// TIA Portal project "MT_SLP333D-IOL_v2" (V18)

(* hardware
DEVICE "S71500/ET200MP station_1"  S7-1500 station
   slot 0: "Rail_0"  Rack  6ES7 590-1***0-0AA0
   slot 1: "PLC_1"  CPU 1516-3 PN/DP  6ES7 516-3AN01-0AB0  V2.8
      slot 3: "CPU display_1"  6ES7591-1BA00-0AA0
      slot 32768: "PROFINET interface_1"  X1
         slot 32769: "Port_1"  X1 P1
         slot 32770: "Port_2"  X1 P2
      slot 33024: "PROFINET interface_2"  X2
         slot 33025: "Port_1"  X2 P1
      slot 33280: "DP interface_1"  X3
      slot 34817: "Virtual CP interface port_1"  Virtual CP interface port  Virtual CP interface port
DEVICE "GSD device_1"  GSD.Device.PN
   slot 0: "Rack"  Rack  V1.0
   slot 0: "bnixg35080b5r067"  BNI XG3-508-0B5-R067  BNI00L3  V1.4.0
      slot 0: "BNI XG3-508-0B5-R067"  BNI XG3-508-0B5-R067
      slot 1: "PN-IO"  PN-IO
         slot 1: "Port XF1"  Port XF1
         slot 2: "Port XF2"  Port XF2
   slot 1: "IO-Link I/O Ports_1"  IO-Link I/O Ports
      slot 0: "BALLUFF 8 Port IO-Link Master"  BALLUFF 8 Port IO-Link Master
   slot 1: "Port deactivated"  Port deactivated
   slot 2: "Port deactivated_1"  Port deactivated
   slot 3: "Port deactivated_2"  Port deactivated
   slot 4: "SLP333D-IOL_Port4I"  IOL_I/O_08/08_Byte + PQI
   slot 5: "Port deactivated_4"  Port deactivated
   slot 6: "Port deactivated_5"  Port deactivated
   slot 7: "Port deactivated_6"  Port deactivated
   slot 8: "Port deactivated_7"  Port deactivated
*)

// ===== PLC "PLC_1"  CPU 1516-3 PN/DP =====

VAR_GLOBAL   // PLC tag table "Default tag table"
   "FirstScan" AT %M1.0 : Bool;
   "SLP/SWP33x_In_Octet0_3" AT %ID1 : DWord;
   "SLP/SWP33x_In_Octet4" AT %IB5 : Byte;
   "SLP/SWP33x_In_Octet5" AT %IB6 : Byte;
   "SLP/SWP33x_In_Octet6" AT %IB7 : Byte;
   "CurrentWeight" AT %MD68 : Real;
   "LowerThreshold" AT %MW72 : UInt;
   "AcyclicCommandIndex" AT %MW74 : UInt;
   "Write_LowerTreshold" AT %M76.0 : Bool;
   "Read_SensorStatus" AT %M76.1 : Bool;
   "Read_AcyclicCommand" AT %M76.2 : Bool;
   "Read_LowerTreshold" AT %M76.3 : Bool;
   "Send_System_Command" AT %M76.4 : Bool;
   "SystemCommand" AT %MW78 : UInt;
   "AcyclicCommandSubindex" AT %MW80 : UInt;
   "AcyclicCommandLength" AT %MW82 : UInt;
   "SensorStatus_SensorNr" AT %MW84 : UInt;
   "Reset_Acyclic_Block" AT %M86.0 : Bool;
   "Smart5Lvl2" AT %M86.1 : Bool;
   "Smart5Lvl3" AT %M86.2 : Bool;
   "Smart5Lvl4" AT %M86.3 : Bool;
   "Smart5Lvl5" AT %M86.4 : Bool;
   "LowerLvlAlarm" AT %M86.5 : Bool;
   "UpperLvlAlarm" AT %M86.6 : Bool;
   "Heartbeat" AT %M86.7 : Bool;
   "CurrentWeightPercent" AT %MD87 : Real;
   "SLP/SWP33x_In_Octet7" AT %IB8 : Byte;
   "SLP/SWP33x_Out_Octet0_3" AT %QD1 : DWord;
   "SLP/SWP33x_Out_Octet6_7" AT %QW7 : Int;
   "ResetCommand" AT %M0.0 : Bool;
   "CommandValue" AT %MD10 : Real;
   "Command" AT %MW15 : Int;
   "WeightMode" AT %MW18 : Int;
   "ProcessType" AT %MW20 : Int;
   "ProcessStatus" AT %MW22 : Int;
   "Write_CommandWithParameter" AT %M76.5 : Bool;
   "ParameterValue" AT %MW91 : UInt;
END_VAR

TYPE "SAI_MB_DeviceStatus"
VERSION : 0.1
   STRUCT
      "Number of Sensors bit 1" : Byte;
      "System Status bit 1" : Bool;
      "System Status bit 2" : Bool;
      "System Status bit 3" : Bool;
      "System Status bit 4" : Bool;
   END_STRUCT;
END_TYPE

TYPE "SAI_SB_3rdStatus"
   STRUCT
      "Measure Unit bit 1" : Bool;
      "Measure Unit bit 2" : Bool;
      "Measure Unit bit 3" : Bool;
      "Measure Unit bit 4" : Bool;
      "Measure Type bit 1" : Bool;
      "Measure Type bit 2" : Bool;
      "Lower Alarm Status" : Bool;
      "Upper Alarm Status" : Bool;
   END_STRUCT;
END_TYPE

TYPE "SAI_SB_2ndStatus"
   STRUCT
      "Smart5 level 5" : Bool;
      "Smart5 level 4" : Bool;
      "Smart5 level 3" : Bool;
      "Smart5 level 2" : Bool;
      Hearbeat : Bool;
   END_STRUCT;
END_TYPE

DATA_BLOCK "SLP/SWP331_IOL_DB"   // DB1
{ S7_Optimized_Access := 'TRUE' }
VERSION : 0.1
// stored: InstanceOfName SLP/SWP331_IOL
"SLP/SWP331_IOL"
BEGIN
END_DATA_BLOCK

DATA_BLOCK "IO_LINK_DEVICE_DB"   // DB2
{ S7_Optimized_Access := 'TRUE' }
AUTHOR : SUP_FA
FAMILY : IO-Link
VERSION : 3.0
// stored: InstanceOfName IO_LINK_DEVICE
"IO_LINK_DEVICE"
BEGIN
END_DATA_BLOCK

DATA_BLOCK "SLP/SWP331_IOL_Acyclic_Commands_DB"   // DB3
{ S7_Optimized_Access := 'TRUE' }
VERSION : 0.1
// stored: InstanceOfName SLP/SWP331_IOL_Acyclic_Commands
"SLP/SWP331_IOL_Acyclic_Commands"
BEGIN
END_DATA_BLOCK

DATA_BLOCK "Data_block_IOL"   // DB14
{ S7_Optimized_Access := 'TRUE' }
VERSION : 0.1
   VAR
      Data : Array[0..231] of Byte;
   END_VAR
BEGIN
END_DATA_BLOCK

FUNCTION_BLOCK "SLP/SWP331_IOL"   // FB1, LAD
{ S7_Optimized_Access := 'TRUE' }
VERSION : 0.1
   VAR_INPUT
      "IO-Link_DevicePort" : Int;
      In_Byte0_3_DWord : DWord;
      In_Byte04 : Byte;
      In_Byte05 : Byte;
      In_Byte06 : Byte;
      In_Byte07 : Byte;
   END_VAR
   VAR_OUTPUT
      CurrentWeight : Real;
      WeightType : String;
      WeightUnit : String;
      Data_OK : Bool;
      Center_Of_Zero : Bool;
      Motion : Bool;
      Net_Mode : Bool;
      Status_Smart5_Lvl_2 : Bool;
      Status_Smart5_Lvl_3 : Bool;
      Status_Smart5_Lvl_4 : Bool;
      Status_Smart5_Lvl_5 : Bool;
      Status_HeartBeat : Bool;
      "Factory adjustment active" : Bool;
      "Last Adjustment Status" : Bool;
      ProcessType : String;
      ProcessType_1 : Int;
      NewWeightUpdate : Bool;
      ProcessStatus : String;
      ProcessStatus_1 : Int;
      Out_Byte0_3_DWord : DWord;
      Out_Byte06_7_Int : Int;
   END_VAR
   VAR_IN_OUT
      "Command Value" : Real;
      Command : Int;
   END_VAR
   VAR
      MeasuredWeightType : Byte;
      MeasuredUnit : Byte;
      ProcessTypeParsen : Byte;
      ProcessStatusParsen : Byte;
      CommandExec : Bool;
   END_VAR
BEGIN

REGION Network 1: Assign IO-Link Device Port Number on the IO-Link Master
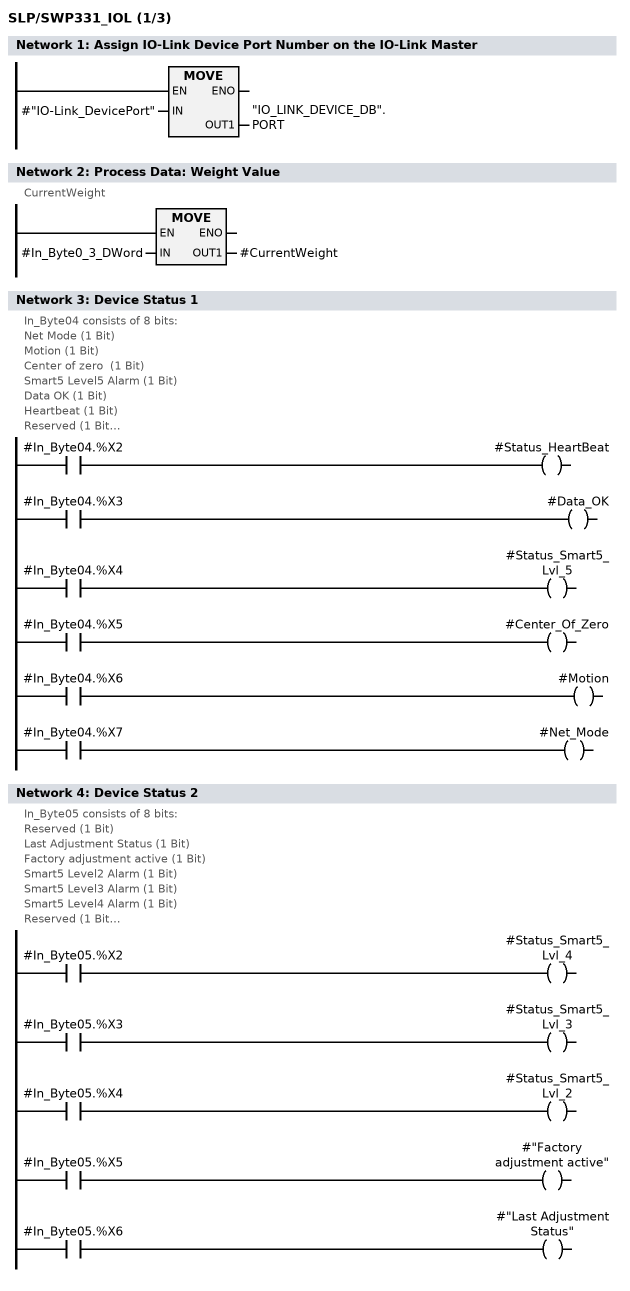
   RUNG wire#powerrail
      Move(in := #"IO-Link_DevicePort", out1 => "IO_LINK_DEVICE_DB".PORT)
   END_RUNG
   // the same network as SCL:
   "IO_LINK_DEVICE_DB".PORT := #"IO-Link_DevicePort";
END_REGION

REGION Network 2: Process Data: Weight Value
   // CurrentWeight
   RUNG wire#powerrail
      Move(in := #In_Byte0_3_DWord, out1 => #CurrentWeight)
   END_RUNG
   // the same network as SCL:
   #CurrentWeight := #In_Byte0_3_DWord;
END_REGION

REGION Network 3: Device Status 1
   // In_Byte04 consists of 8 bits:
   // 
   // Net Mode (1 Bit) 
   // Motion (1 Bit) 
   // Center of zero  (1 Bit) 
   // Smart5 Level5 Alarm (1 Bit) 
   // Data OK (1 Bit) 
   // Heartbeat (1 Bit) 
   // Reserved (1 Bit) 
   // Reserved (1 Bit)
   RUNG wire#powerrail
      Contact( #In_Byte04.%X2 )
      Coil( #Status_HeartBeat )
   END_RUNG
   RUNG wire#powerrail
      Contact( #In_Byte04.%X3 )
      Coil( #Data_OK )
   END_RUNG
   RUNG wire#powerrail
      Contact( #In_Byte04.%X4 )
      Coil( #Status_Smart5_Lvl_5 )
   END_RUNG
   RUNG wire#powerrail
      Contact( #In_Byte04.%X5 )
      Coil( #Center_Of_Zero )
   END_RUNG
   RUNG wire#powerrail
      Contact( #In_Byte04.%X6 )
      Coil( #Motion )
   END_RUNG
   RUNG wire#powerrail
      Contact( #In_Byte04.%X7 )
      Coil( #Net_Mode )
   END_RUNG
   // the same network as SCL:
   #Status_HeartBeat := #In_Byte04.%X2;
   #Data_OK := #In_Byte04.%X3;
   #Status_Smart5_Lvl_5 := #In_Byte04.%X4;
   #Center_Of_Zero := #In_Byte04.%X5;
   #Motion := #In_Byte04.%X6;
   #Net_Mode := #In_Byte04.%X7;
END_REGION

REGION Network 4: Device Status 2
   // In_Byte05 consists of 8 bits:
   // 
   // Reserved (1 Bit) 
   // Last Adjustment Status (1 Bit) 
   // Factory adjustment active (1 Bit) 
   // Smart5 Level2 Alarm (1 Bit)
   // Smart5 Level3 Alarm (1 Bit) 
   // Smart5 Level4 Alarm (1 Bit) 
   // Reserved (1 Bit) 
   // Reserved (1 Bit)
   RUNG wire#powerrail
      Contact( #In_Byte05.%X2 )
      Coil( #Status_Smart5_Lvl_4 )
   END_RUNG
   RUNG wire#powerrail
      Contact( #In_Byte05.%X3 )
      Coil( #Status_Smart5_Lvl_3 )
   END_RUNG
   RUNG wire#powerrail
      Contact( #In_Byte05.%X4 )
      Coil( #Status_Smart5_Lvl_2 )
   END_RUNG
   RUNG wire#powerrail
      Contact( #In_Byte05.%X5 )
      Coil( #"Factory adjustment active" )
   END_RUNG
   RUNG wire#powerrail
      Contact( #In_Byte05.%X6 )
      Coil( #"Last Adjustment Status" )
   END_RUNG
   // the same network as SCL:
   #Status_Smart5_Lvl_4 := #In_Byte05.%X2;
   #Status_Smart5_Lvl_3 := #In_Byte05.%X3;
   #Status_Smart5_Lvl_2 := #In_Byte05.%X4;
   #"Factory adjustment active" := #In_Byte05.%X5;
   #"Last Adjustment Status" := #In_Byte05.%X6;
END_REGION

REGION Network 5: Device Status 3
   // In_Byte06 consists of 8 bits:
   // 
   // Process Type (3 Bit) 
   // New weight update (1 Bit) 
   // Process Status (4 Bit)
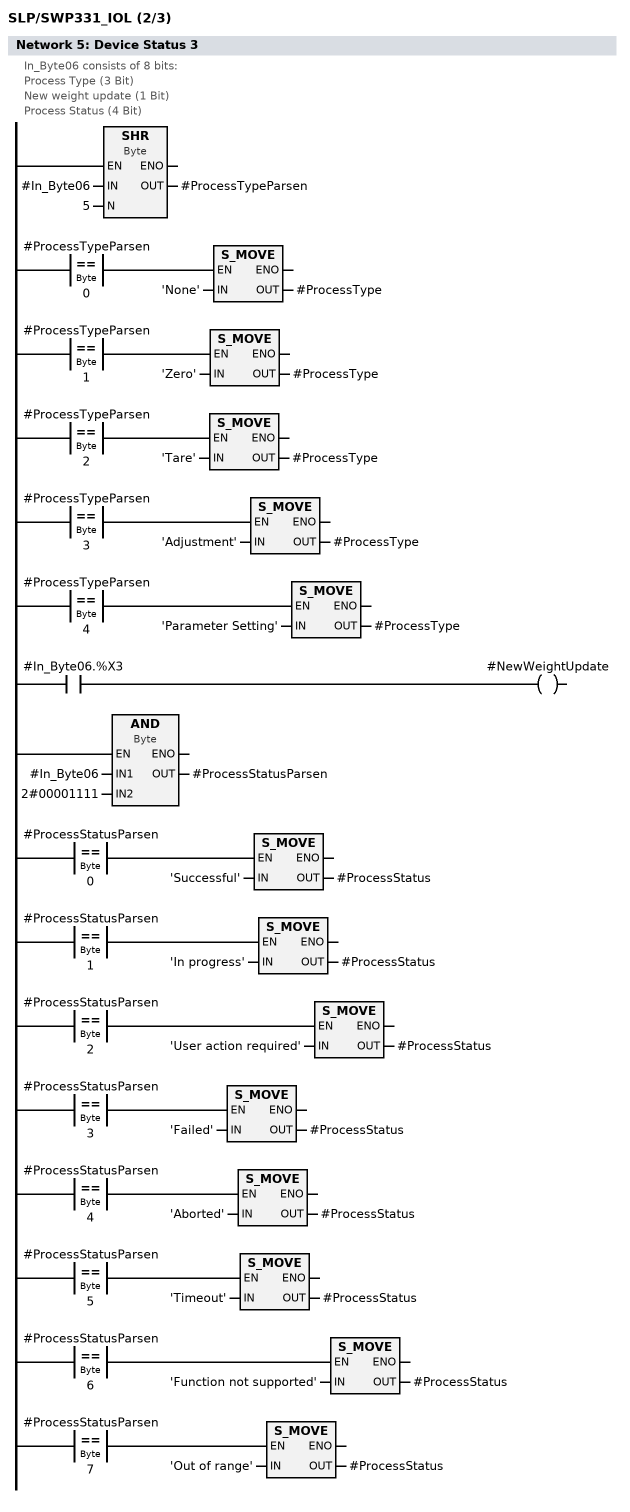
   RUNG wire#powerrail
      { S7_Templates := "SrcType := Byte" } Shr(in := #In_Byte06, n := 5, out => #ProcessTypeParsen)
   END_RUNG
   RUNG wire#powerrail
      { S7_Templates := "SrcType := Byte" } EQ_Contact(in1 := #ProcessTypeParsen, in2 := 0)
      S_Move(in := 'None', out => #ProcessType)
   END_RUNG
   RUNG wire#powerrail
      { S7_Templates := "SrcType := Byte" } EQ_Contact(in1 := #ProcessTypeParsen, in2 := 1)
      S_Move(in := 'Zero', out => #ProcessType)
   END_RUNG
   RUNG wire#powerrail
      { S7_Templates := "SrcType := Byte" } EQ_Contact(in1 := #ProcessTypeParsen, in2 := 2)
      S_Move(in := 'Tare', out => #ProcessType)
   END_RUNG
   RUNG wire#powerrail
      { S7_Templates := "SrcType := Byte" } EQ_Contact(in1 := #ProcessTypeParsen, in2 := 3)
      S_Move(in := 'Adjustment', out => #ProcessType)
   END_RUNG
   RUNG wire#powerrail
      { S7_Templates := "SrcType := Byte" } EQ_Contact(in1 := #ProcessTypeParsen, in2 := 4)
      S_Move(in := 'Parameter Setting', out => #ProcessType)
   END_RUNG
   RUNG wire#powerrail
      Contact( #In_Byte06.%X3 )
      Coil( #NewWeightUpdate )
   END_RUNG
   RUNG wire#powerrail
      { S7_Templates := "SrcType := Byte" } And(in1 := #In_Byte06, in2 := 2#00001111, out => #ProcessStatusParsen)
   END_RUNG
   RUNG wire#powerrail
      { S7_Templates := "SrcType := Byte" } EQ_Contact(in1 := #ProcessStatusParsen, in2 := 0)
      S_Move(in := 'Successful', out => #ProcessStatus)
   END_RUNG
   RUNG wire#powerrail
      { S7_Templates := "SrcType := Byte" } EQ_Contact(in1 := #ProcessStatusParsen, in2 := 1)
      S_Move(in := 'In progress', out => #ProcessStatus)
   END_RUNG
   RUNG wire#powerrail
      { S7_Templates := "SrcType := Byte" } EQ_Contact(in1 := #ProcessStatusParsen, in2 := 2)
      S_Move(in := 'User action required', out => #ProcessStatus)
   END_RUNG
   RUNG wire#powerrail
      { S7_Templates := "SrcType := Byte" } EQ_Contact(in1 := #ProcessStatusParsen, in2 := 3)
      S_Move(in := 'Failed', out => #ProcessStatus)
   END_RUNG
   RUNG wire#powerrail
      { S7_Templates := "SrcType := Byte" } EQ_Contact(in1 := #ProcessStatusParsen, in2 := 4)
      S_Move(in := 'Aborted', out => #ProcessStatus)
   END_RUNG
   RUNG wire#powerrail
      { S7_Templates := "SrcType := Byte" } EQ_Contact(in1 := #ProcessStatusParsen, in2 := 5)
      S_Move(in := 'Timeout', out => #ProcessStatus)
   END_RUNG
   RUNG wire#powerrail
      { S7_Templates := "SrcType := Byte" } EQ_Contact(in1 := #ProcessStatusParsen, in2 := 6)
      S_Move(in := 'Function not supported', out => #ProcessStatus)
   END_RUNG
   RUNG wire#powerrail
      { S7_Templates := "SrcType := Byte" } EQ_Contact(in1 := #ProcessStatusParsen, in2 := 7)
      S_Move(in := 'Out of range', out => #ProcessStatus)
   END_RUNG
   // the same network as SCL:
   #ProcessTypeParsen := SHR(IN := #In_Byte06, N := 5);
   IF #ProcessTypeParsen = 0 THEN #ProcessType := 'None'; END_IF;
   IF #ProcessTypeParsen = 1 THEN #ProcessType := 'Zero'; END_IF;
   IF #ProcessTypeParsen = 2 THEN #ProcessType := 'Tare'; END_IF;
   IF #ProcessTypeParsen = 3 THEN #ProcessType := 'Adjustment'; END_IF;
   IF #ProcessTypeParsen = 4 THEN #ProcessType := 'Parameter Setting'; END_IF;
   #NewWeightUpdate := #In_Byte06.%X3;
   #ProcessStatusParsen := #In_Byte06 AND 2#00001111;
   IF #ProcessStatusParsen = 0 THEN #ProcessStatus := 'Successful'; END_IF;
   IF #ProcessStatusParsen = 1 THEN #ProcessStatus := 'In progress'; END_IF;
   IF #ProcessStatusParsen = 2 THEN #ProcessStatus := 'User action required'; END_IF;
   IF #ProcessStatusParsen = 3 THEN #ProcessStatus := 'Failed'; END_IF;
   IF #ProcessStatusParsen = 4 THEN #ProcessStatus := 'Aborted'; END_IF;
   IF #ProcessStatusParsen = 5 THEN #ProcessStatus := 'Timeout'; END_IF;
   IF #ProcessStatusParsen = 6 THEN #ProcessStatus := 'Function not supported'; END_IF;
   IF #ProcessStatusParsen = 7 THEN #ProcessStatus := 'Out of range'; END_IF;
END_REGION

REGION Network 6: Weight Information
   // In_Byte07 consists of 8 bits:
   // Weight Type (4 Bits)
   // Weight Unit (4 Bits)
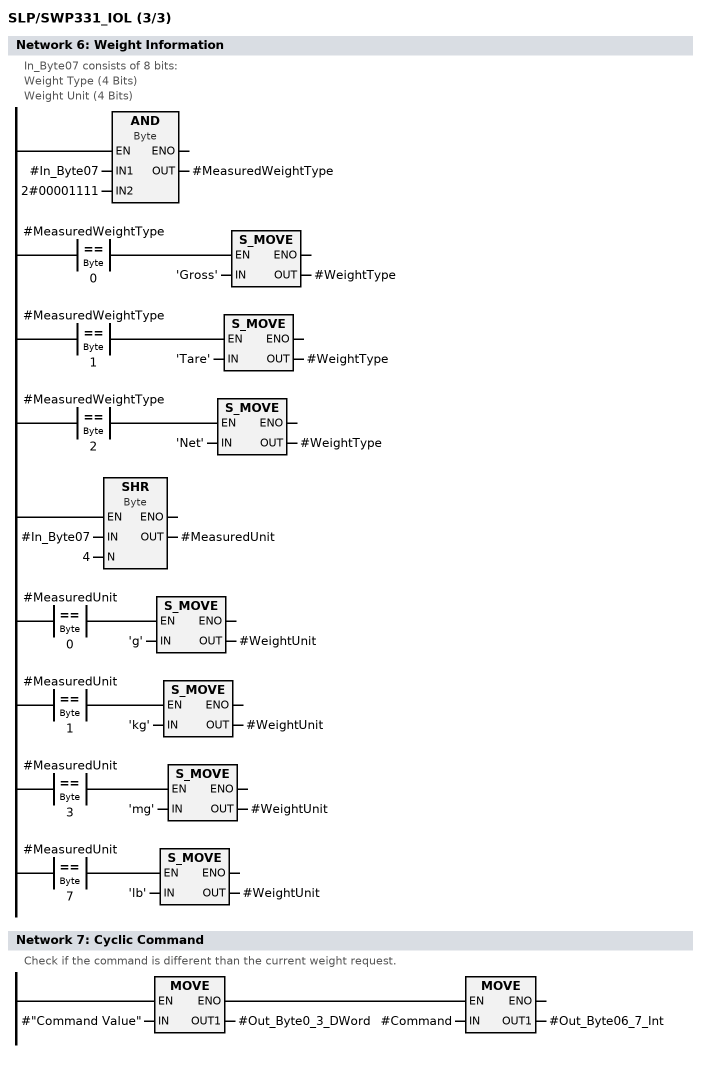
   RUNG wire#powerrail
      { S7_Templates := "SrcType := Byte" } And(in1 := #In_Byte07, in2 := 2#00001111, out => #MeasuredWeightType)
   END_RUNG
   RUNG wire#powerrail
      { S7_Templates := "SrcType := Byte" } EQ_Contact(in1 := #MeasuredWeightType, in2 := 0)
      S_Move(in := 'Gross', out => #WeightType)
   END_RUNG
   RUNG wire#powerrail
      { S7_Templates := "SrcType := Byte" } EQ_Contact(in1 := #MeasuredWeightType, in2 := 1)
      S_Move(in := 'Tare', out => #WeightType)
   END_RUNG
   RUNG wire#powerrail
      { S7_Templates := "SrcType := Byte" } EQ_Contact(in1 := #MeasuredWeightType, in2 := 2)
      S_Move(in := 'Net', out => #WeightType)
   END_RUNG
   RUNG wire#powerrail
      { S7_Templates := "SrcType := Byte" } Shr(in := #In_Byte07, n := 4, out => #MeasuredUnit)
   END_RUNG
   RUNG wire#powerrail
      { S7_Templates := "SrcType := Byte" } EQ_Contact(in1 := #MeasuredUnit, in2 := 0)
      S_Move(in := 'g', out => #WeightUnit)
   END_RUNG
   RUNG wire#powerrail
      { S7_Templates := "SrcType := Byte" } EQ_Contact(in1 := #MeasuredUnit, in2 := 1)
      S_Move(in := 'kg', out => #WeightUnit)
   END_RUNG
   RUNG wire#powerrail
      { S7_Templates := "SrcType := Byte" } EQ_Contact(in1 := #MeasuredUnit, in2 := 3)
      S_Move(in := 'mg', out => #WeightUnit)
   END_RUNG
   RUNG wire#powerrail
      { S7_Templates := "SrcType := Byte" } EQ_Contact(in1 := #MeasuredUnit, in2 := 7)
      S_Move(in := 'lb', out => #WeightUnit)
   END_RUNG
   // the same network as SCL:
   #MeasuredWeightType := #In_Byte07 AND 2#00001111;
   IF #MeasuredWeightType = 0 THEN #WeightType := 'Gross'; END_IF;
   IF #MeasuredWeightType = 1 THEN #WeightType := 'Tare'; END_IF;
   IF #MeasuredWeightType = 2 THEN #WeightType := 'Net'; END_IF;
   #MeasuredUnit := SHR(IN := #In_Byte07, N := 4);
   IF #MeasuredUnit = 0 THEN #WeightUnit := 'g'; END_IF;
   IF #MeasuredUnit = 1 THEN #WeightUnit := 'kg'; END_IF;
   IF #MeasuredUnit = 3 THEN #WeightUnit := 'mg'; END_IF;
   IF #MeasuredUnit = 7 THEN #WeightUnit := 'lb'; END_IF;
END_REGION

REGION Network 7: Cyclic Command
   // Check if the command is different than the current weight request.
   RUNG wire#powerrail
      Move(in := #"Command Value", out1 => #Out_Byte0_3_DWord)
      Move(in := #Command, out1 => #Out_Byte06_7_Int)
   END_RUNG
   // the same network as SCL:
   #Out_Byte0_3_DWord := #"Command Value";
   #Out_Byte06_7_Int := #Command;
END_REGION
END_FUNCTION_BLOCK

FUNCTION_BLOCK "SLP/SWP331_IOL_Acyclic_Commands"   // FB2, LAD
{ S7_Optimized_Access := 'TRUE' }
VERSION : 0.1
   VAR_INPUT
      SystemCommand : UInt;
      AcyclicCommandIndex : UInt;
      AcyclicCommandSubindex : UInt;
      AcyclicCommandLength : UInt;
      ParameterValue : UInt;
   END_VAR
   VAR_OUTPUT
      SensorStatus : Byte;
      ErrorCode : DWord;
      Done : Bool;
   END_VAR
   VAR_IN_OUT
      Send_SystemCmd : Bool;
      Write_AcyclicCommandWithParameter : Bool;
      Read_AcyclicCommand : Bool;
      ResetAcyclicBlock : Bool;
   END_VAR
   VAR
      WriteStep : SInt;
      ReadStep : SInt;
      Cmd_RWTrigger : Bool;
   END_VAR
   VAR_TEMP   // added for the SCL form of the ladder/FBD networks
      _w1 : Bool;
      _w2 : Bool;
      _w3 : Bool;
      _w4 : Bool;
      _w5 : Bool;
      _w6 : Bool;
   END_VAR
BEGIN

REGION Network 1: Send Acyclic Command
   // Change the variable #SystemCommand in the Application Block and trigger the #Send_SystemCmd to send a system command to the device.
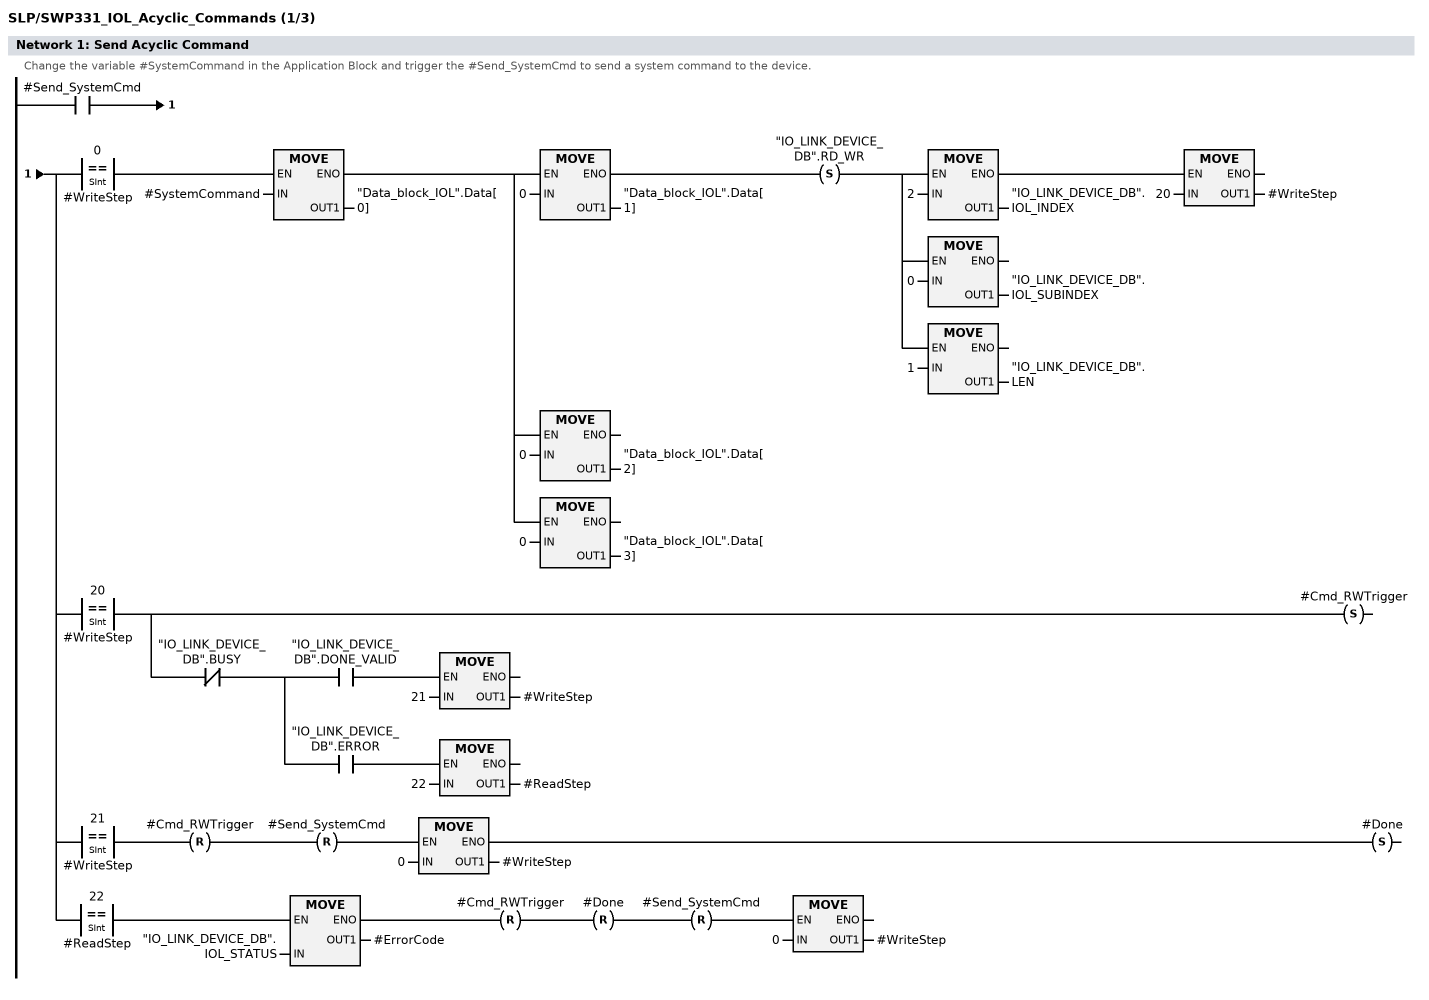
   RUNG wire#powerrail
      Contact( #Send_SystemCmd )
      wire#w1
      { S7_Templates := "SrcType := SInt" } EQ_Contact(in1 := 0, in2 := #WriteStep)
      Move(in := #SystemCommand, out1 => "Data_block_IOL".Data[0])
      wire#w2
      Move(in := 0, out1 => "Data_block_IOL".Data[1])
      S_Coil( "IO_LINK_DEVICE_DB".RD_WR )
      wire#w3
      Move(in := 2, out1 => "IO_LINK_DEVICE_DB".IOL_INDEX)
      Move(in := 20, out1 => #WriteStep)
   END_RUNG
   RUNG wire#w3
      Move(in := 0, out1 => "IO_LINK_DEVICE_DB".IOL_SUBINDEX)
   END_RUNG
   RUNG wire#w3
      Move(in := 1, out1 => "IO_LINK_DEVICE_DB".LEN)
   END_RUNG
   RUNG wire#w2
      Move(in := 0, out1 => "Data_block_IOL".Data[2])
   END_RUNG
   RUNG wire#w2
      Move(in := 0, out1 => "Data_block_IOL".Data[3])
   END_RUNG
   RUNG wire#w1
      { S7_Templates := "SrcType := SInt" } EQ_Contact(in1 := 20, in2 := #WriteStep)
      wire#w4
      S_Coil( #Cmd_RWTrigger )
   END_RUNG
   RUNG wire#w4
      I_Contact( "IO_LINK_DEVICE_DB".BUSY )
      wire#w5
      Contact( "IO_LINK_DEVICE_DB".DONE_VALID )
      Move(in := 21, out1 => #WriteStep)
   END_RUNG
   RUNG wire#w5
      Contact( "IO_LINK_DEVICE_DB".ERROR )
      Move(in := 22, out1 => #ReadStep)
   END_RUNG
   RUNG wire#w1
      { S7_Templates := "SrcType := SInt" } EQ_Contact(in1 := 21, in2 := #WriteStep)
      R_Coil( #Cmd_RWTrigger )
      R_Coil( #Send_SystemCmd )
      Move(in := 0, out1 => #WriteStep)
      S_Coil( #Done )
   END_RUNG
   RUNG wire#w1
      { S7_Templates := "SrcType := SInt" } EQ_Contact(in1 := 22, in2 := #ReadStep)
      Move(in := "IO_LINK_DEVICE_DB".IOL_STATUS, out1 => #ErrorCode)
      R_Coil( #Cmd_RWTrigger )
      R_Coil( #Done )
      R_Coil( #Send_SystemCmd )
      Move(in := 0, out1 => #WriteStep)
   END_RUNG
   // the same network as SCL:
   IF #Send_SystemCmd AND (0 = #WriteStep) THEN
       "Data_block_IOL".Data[0] := #SystemCommand;
       "Data_block_IOL".Data[1] := 0;
       "IO_LINK_DEVICE_DB".RD_WR := TRUE;
       "IO_LINK_DEVICE_DB".IOL_INDEX := 2;
   END_IF;
   #_w1 := #Send_SystemCmd AND (0 = #WriteStep);
   #_w2 := #Send_SystemCmd AND (0 = #WriteStep);
   IF #_w2 THEN
       #WriteStep := 20;
       "IO_LINK_DEVICE_DB".IOL_SUBINDEX := 0;
       "IO_LINK_DEVICE_DB".LEN := 1;
   END_IF;
   IF #_w1 THEN
       "Data_block_IOL".Data[2] := 0;
       "Data_block_IOL".Data[3] := 0;
   END_IF;
   #_w3 := #Send_SystemCmd AND (20 = #WriteStep);
   IF #_w3 THEN #Cmd_RWTrigger := TRUE; END_IF;
   #_w4 := #_w3 AND NOT "IO_LINK_DEVICE_DB".BUSY;
   IF #_w4 AND "IO_LINK_DEVICE_DB".DONE_VALID THEN #WriteStep := 21; END_IF;
   IF #_w4 AND "IO_LINK_DEVICE_DB".ERROR THEN #ReadStep := 22; END_IF;
   IF #Send_SystemCmd AND (21 = #WriteStep) THEN #Cmd_RWTrigger := FALSE; END_IF;
   #_w5 := #Send_SystemCmd AND (21 = #WriteStep);
   #_w6 := #Send_SystemCmd;
   IF #_w5 THEN
       #Send_SystemCmd := FALSE;
       #WriteStep := 0;
       #Done := TRUE;
   END_IF;
   IF #_w6 AND (22 = #ReadStep) THEN
       #ErrorCode := "IO_LINK_DEVICE_DB".IOL_STATUS;
       #Cmd_RWTrigger := FALSE;
       #Done := FALSE;
       #Send_SystemCmd := FALSE;
       #WriteStep := 0;
   END_IF;
END_REGION

REGION Network 2: Read Acyclic Command
   // Change the variables value #AcyclicCommandIndex, #AcyclicCommandSubindex and #AcyclicCommandLength in the Application Block and trigger the #Read_AcyclicCommand to send an acyclic command to the device.
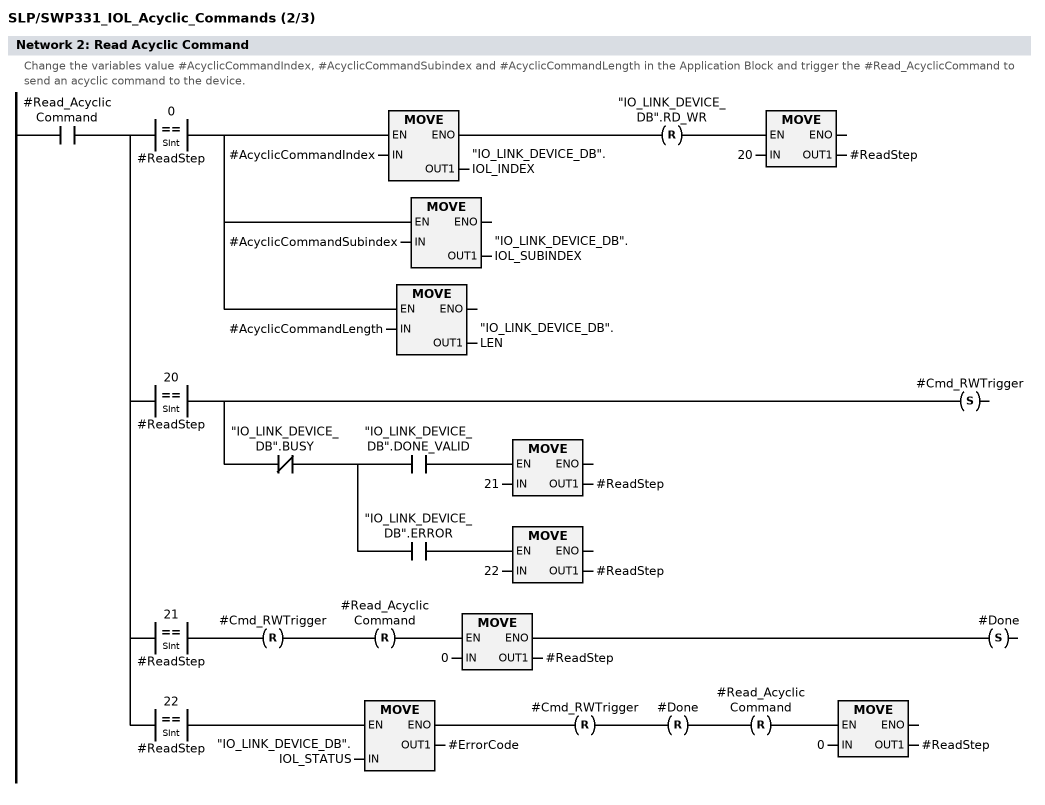
   RUNG wire#powerrail
      Contact( #Read_AcyclicCommand )
      wire#w1
      { S7_Templates := "SrcType := SInt" } EQ_Contact(in1 := 0, in2 := #ReadStep)
      wire#w2
      Move(in := #AcyclicCommandIndex, out1 => "IO_LINK_DEVICE_DB".IOL_INDEX)
      R_Coil( "IO_LINK_DEVICE_DB".RD_WR )
      Move(in := 20, out1 => #ReadStep)
   END_RUNG
   RUNG wire#w2
      Move(in := #AcyclicCommandSubindex, out1 => "IO_LINK_DEVICE_DB".IOL_SUBINDEX)
   END_RUNG
   RUNG wire#w2
      Move(in := #AcyclicCommandLength, out1 => "IO_LINK_DEVICE_DB".LEN)
   END_RUNG
   RUNG wire#w1
      { S7_Templates := "SrcType := SInt" } EQ_Contact(in1 := 20, in2 := #ReadStep)
      wire#w3
      S_Coil( #Cmd_RWTrigger )
   END_RUNG
   RUNG wire#w3
      I_Contact( "IO_LINK_DEVICE_DB".BUSY )
      wire#w4
      Contact( "IO_LINK_DEVICE_DB".DONE_VALID )
      Move(in := 21, out1 => #ReadStep)
   END_RUNG
   RUNG wire#w4
      Contact( "IO_LINK_DEVICE_DB".ERROR )
      Move(in := 22, out1 => #ReadStep)
   END_RUNG
   RUNG wire#w1
      { S7_Templates := "SrcType := SInt" } EQ_Contact(in1 := 21, in2 := #ReadStep)
      R_Coil( #Cmd_RWTrigger )
      R_Coil( #Read_AcyclicCommand )
      Move(in := 0, out1 => #ReadStep)
      S_Coil( #Done )
   END_RUNG
   RUNG wire#w1
      { S7_Templates := "SrcType := SInt" } EQ_Contact(in1 := 22, in2 := #ReadStep)
      Move(in := "IO_LINK_DEVICE_DB".IOL_STATUS, out1 => #ErrorCode)
      R_Coil( #Cmd_RWTrigger )
      R_Coil( #Done )
      R_Coil( #Read_AcyclicCommand )
      Move(in := 0, out1 => #ReadStep)
   END_RUNG
   // the same network as SCL:
   IF #Read_AcyclicCommand AND (0 = #ReadStep) THEN
       "IO_LINK_DEVICE_DB".IOL_INDEX := #AcyclicCommandIndex;
       "IO_LINK_DEVICE_DB".RD_WR := FALSE;
   END_IF;
   #_w1 := #Read_AcyclicCommand AND (0 = #ReadStep);
   IF #_w1 THEN
       #ReadStep := 20;
       "IO_LINK_DEVICE_DB".IOL_SUBINDEX := #AcyclicCommandSubindex;
       "IO_LINK_DEVICE_DB".LEN := #AcyclicCommandLength;
   END_IF;
   #_w2 := #Read_AcyclicCommand AND (20 = #ReadStep);
   IF #_w2 THEN #Cmd_RWTrigger := TRUE; END_IF;
   #_w3 := #_w2 AND NOT "IO_LINK_DEVICE_DB".BUSY;
   IF #_w3 AND "IO_LINK_DEVICE_DB".DONE_VALID THEN #ReadStep := 21; END_IF;
   IF #_w3 AND "IO_LINK_DEVICE_DB".ERROR THEN #ReadStep := 22; END_IF;
   IF #Read_AcyclicCommand AND (21 = #ReadStep) THEN #Cmd_RWTrigger := FALSE; END_IF;
   #_w4 := #Read_AcyclicCommand AND (21 = #ReadStep);
   #_w5 := #Read_AcyclicCommand;
   IF #_w4 THEN
       #Read_AcyclicCommand := FALSE;
       #ReadStep := 0;
       #Done := TRUE;
   END_IF;
   IF #_w5 AND (22 = #ReadStep) THEN
       #ErrorCode := "IO_LINK_DEVICE_DB".IOL_STATUS;
       #Cmd_RWTrigger := FALSE;
       #Done := FALSE;
       #Read_AcyclicCommand := FALSE;
       #ReadStep := 0;
   END_IF;
END_REGION

REGION Network 3: Write Acyclic Command
   // Change the variables value #AcyclicCommandIndex, #AcyclicCommandSubindex #ParameterValue and #AcyclicCommandLength in the Application Block and trigger the #Write_AcyclicCommand to send an acyclic command to the device.
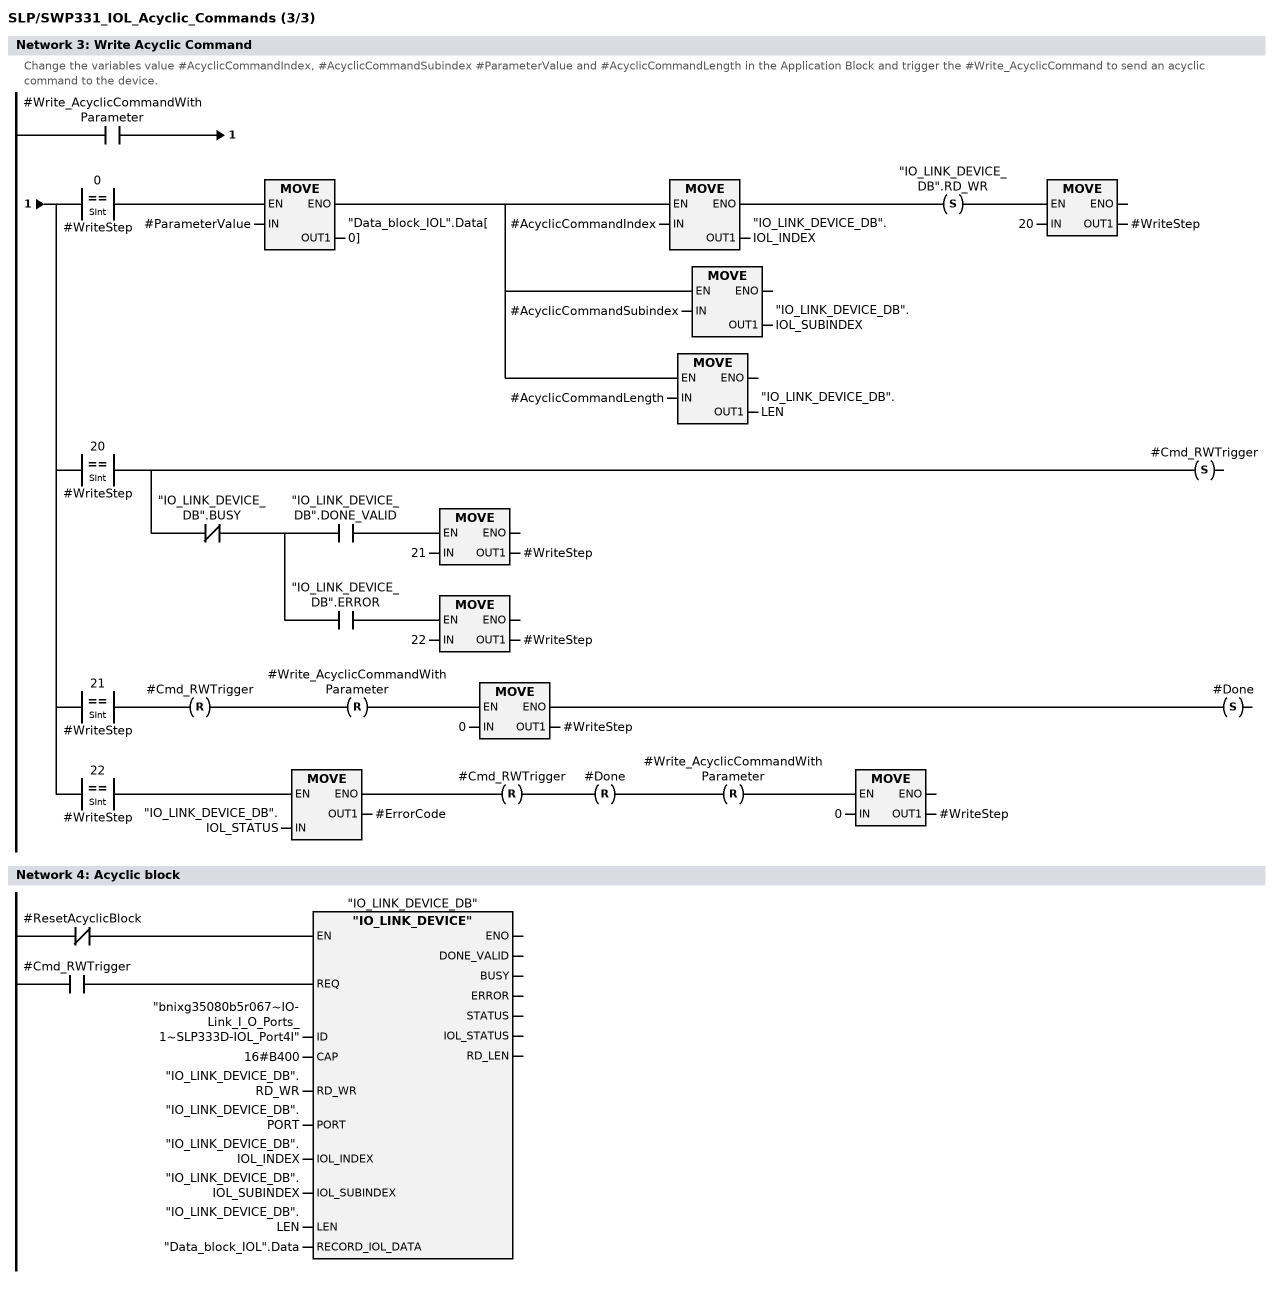
   RUNG wire#powerrail
      Contact( #Write_AcyclicCommandWithParameter )
      wire#w1
      { S7_Templates := "SrcType := SInt" } EQ_Contact(in1 := 0, in2 := #WriteStep)
      Move(in := #ParameterValue, out1 => "Data_block_IOL".Data[0])
      wire#w2
      Move(in := #AcyclicCommandIndex, out1 => "IO_LINK_DEVICE_DB".IOL_INDEX)
      S_Coil( "IO_LINK_DEVICE_DB".RD_WR )
      Move(in := 20, out1 => #WriteStep)
   END_RUNG
   RUNG wire#w2
      Move(in := #AcyclicCommandSubindex, out1 => "IO_LINK_DEVICE_DB".IOL_SUBINDEX)
   END_RUNG
   RUNG wire#w2
      Move(in := #AcyclicCommandLength, out1 => "IO_LINK_DEVICE_DB".LEN)
   END_RUNG
   RUNG wire#w1
      { S7_Templates := "SrcType := SInt" } EQ_Contact(in1 := 20, in2 := #WriteStep)
      wire#w3
      S_Coil( #Cmd_RWTrigger )
   END_RUNG
   RUNG wire#w3
      I_Contact( "IO_LINK_DEVICE_DB".BUSY )
      wire#w4
      Contact( "IO_LINK_DEVICE_DB".DONE_VALID )
      Move(in := 21, out1 => #WriteStep)
   END_RUNG
   RUNG wire#w4
      Contact( "IO_LINK_DEVICE_DB".ERROR )
      Move(in := 22, out1 => #WriteStep)
   END_RUNG
   RUNG wire#w1
      { S7_Templates := "SrcType := SInt" } EQ_Contact(in1 := 21, in2 := #WriteStep)
      R_Coil( #Cmd_RWTrigger )
      R_Coil( #Write_AcyclicCommandWithParameter )
      Move(in := 0, out1 => #WriteStep)
      S_Coil( #Done )
   END_RUNG
   RUNG wire#w1
      { S7_Templates := "SrcType := SInt" } EQ_Contact(in1 := 22, in2 := #WriteStep)
      Move(in := "IO_LINK_DEVICE_DB".IOL_STATUS, out1 => #ErrorCode)
      R_Coil( #Cmd_RWTrigger )
      R_Coil( #Done )
      R_Coil( #Write_AcyclicCommandWithParameter )
      Move(in := 0, out1 => #WriteStep)
   END_RUNG
   // the same network as SCL:
   IF #Write_AcyclicCommandWithParameter AND (0 = #WriteStep) THEN
       "Data_block_IOL".Data[0] := #ParameterValue;
       "IO_LINK_DEVICE_DB".IOL_INDEX := #AcyclicCommandIndex;
       "IO_LINK_DEVICE_DB".RD_WR := TRUE;
   END_IF;
   #_w1 := #Write_AcyclicCommandWithParameter AND (0 = #WriteStep);
   IF #_w1 THEN
       #WriteStep := 20;
       "IO_LINK_DEVICE_DB".IOL_SUBINDEX := #AcyclicCommandSubindex;
       "IO_LINK_DEVICE_DB".LEN := #AcyclicCommandLength;
   END_IF;
   #_w2 := #Write_AcyclicCommandWithParameter AND (20 = #WriteStep);
   IF #_w2 THEN #Cmd_RWTrigger := TRUE; END_IF;
   #_w3 := #_w2 AND NOT "IO_LINK_DEVICE_DB".BUSY;
   IF #_w3 AND "IO_LINK_DEVICE_DB".DONE_VALID THEN #WriteStep := 21; END_IF;
   IF #_w3 AND "IO_LINK_DEVICE_DB".ERROR THEN #WriteStep := 22; END_IF;
   IF #Write_AcyclicCommandWithParameter AND (21 = #WriteStep) THEN #Cmd_RWTrigger := FALSE; END_IF;
   #_w4 := #Write_AcyclicCommandWithParameter AND (21 = #WriteStep);
   #_w5 := #Write_AcyclicCommandWithParameter;
   IF #_w4 THEN
       #Write_AcyclicCommandWithParameter := FALSE;
       #WriteStep := 0;
       #Done := TRUE;
   END_IF;
   IF #_w5 AND (22 = #WriteStep) THEN
       #ErrorCode := "IO_LINK_DEVICE_DB".IOL_STATUS;
       #Cmd_RWTrigger := FALSE;
       #Done := FALSE;
       #Write_AcyclicCommandWithParameter := FALSE;
       #WriteStep := 0;
   END_IF;
END_REGION

REGION Network 4: Acyclic block
   RUNG wire#powerrail
      I_Contact( #ResetAcyclicBlock )
      "IO_LINK_DEVICE_DB"(REQ := wire#w1, ID := "bnixg35080b5r067~IO-Link_I_O_Ports_1~SLP333D-IOL_Port4I", CAP := 16#B400, RD_WR := "IO_LINK_DEVICE_DB".RD_WR, PORT := "IO_LINK_DEVICE_DB".PORT, IOL_INDEX := "IO_LINK_DEVICE_DB".IOL_INDEX, IOL_SUBINDEX := "IO_LINK_DEVICE_DB".IOL_SUBINDEX, LEN := "IO_LINK_DEVICE_DB".LEN, RECORD_IOL_DATA := "Data_block_IOL".Data, DONE_VALID =>, BUSY =>, ERROR =>, STATUS =>, IOL_STATUS =>, RD_LEN =>)
   END_RUNG
   RUNG wire#powerrail
      Contact( #Cmd_RWTrigger )
   END_RUNG wire#w1
   // the same network as SCL:
   IF NOT #ResetAcyclicBlock THEN
       "IO_LINK_DEVICE_DB"(REQ := #Cmd_RWTrigger,   // "IO_LINK_DEVICE"
                           ID := "bnixg35080b5r067~IO-Link_I_O_Ports_1~SLP333D-IOL_Port4I",
                           CAP := 16#B400,
                           RD_WR := "IO_LINK_DEVICE_DB".RD_WR,
                           PORT := "IO_LINK_DEVICE_DB".PORT,
                           IOL_INDEX := "IO_LINK_DEVICE_DB".IOL_INDEX,
                           IOL_SUBINDEX := "IO_LINK_DEVICE_DB".IOL_SUBINDEX,
                           LEN := "IO_LINK_DEVICE_DB".LEN,
                           RECORD_IOL_DATA := "Data_block_IOL".Data);
   END_IF;
END_REGION
END_FUNCTION_BLOCK

FUNCTION "MT_IND_Application" : Void   // FC1, LAD
{ S7_Optimized_Access := 'TRUE' }
VERSION : 0.1
BEGIN

REGION Network 1: Cyclic Data
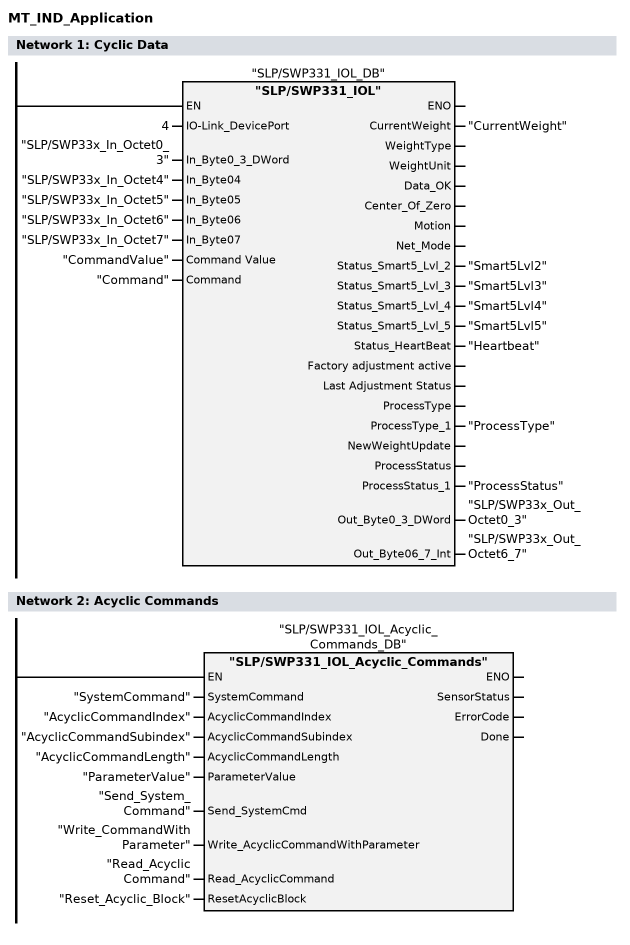
   RUNG wire#powerrail
      "SLP/SWP331_IOL_DB"("IO-Link_DevicePort" := 4, In_Byte0_3_DWord := "SLP/SWP33x_In_Octet0_3", In_Byte04 := "SLP/SWP33x_In_Octet4", In_Byte05 := "SLP/SWP33x_In_Octet5", In_Byte06 := "SLP/SWP33x_In_Octet6", In_Byte07 := "SLP/SWP33x_In_Octet7", "Command Value" := "CommandValue", Command := "Command", CurrentWeight => "CurrentWeight", WeightType =>, WeightUnit =>, Data_OK =>, Center_Of_Zero =>, Motion =>, Net_Mode =>, Status_Smart5_Lvl_2 => "Smart5Lvl2", Status_Smart5_Lvl_3 => "Smart5Lvl3", Status_Smart5_Lvl_4 => "Smart5Lvl4", Status_Smart5_Lvl_5 => "Smart5Lvl5", Status_HeartBeat => "Heartbeat", "Factory adjustment active" =>, "Last Adjustment Status" =>, ProcessType =>, ProcessType_1 => "ProcessType", NewWeightUpdate =>, ProcessStatus =>, ProcessStatus_1 => "ProcessStatus", Out_Byte0_3_DWord => "SLP/SWP33x_Out_Octet0_3", Out_Byte06_7_Int => "SLP/SWP33x_Out_Octet6_7")
   END_RUNG
   // the same network as SCL:
   "SLP/SWP331_IOL_DB"("IO-Link_DevicePort" := 4,   // "SLP/SWP331_IOL"
                       In_Byte0_3_DWord := "SLP/SWP33x_In_Octet0_3",
                       In_Byte04 := "SLP/SWP33x_In_Octet4",
                       In_Byte05 := "SLP/SWP33x_In_Octet5",
                       In_Byte06 := "SLP/SWP33x_In_Octet6",
                       In_Byte07 := "SLP/SWP33x_In_Octet7",
                       "Command Value" := "CommandValue",
                       Command := "Command",
                       CurrentWeight => "CurrentWeight",
                       Status_Smart5_Lvl_2 => "Smart5Lvl2",
                       Status_Smart5_Lvl_3 => "Smart5Lvl3",
                       Status_Smart5_Lvl_4 => "Smart5Lvl4",
                       Status_Smart5_Lvl_5 => "Smart5Lvl5",
                       Status_HeartBeat => "Heartbeat",
                       ProcessType_1 => "ProcessType",
                       ProcessStatus_1 => "ProcessStatus",
                       Out_Byte0_3_DWord => "SLP/SWP33x_Out_Octet0_3",
                       Out_Byte06_7_Int => "SLP/SWP33x_Out_Octet6_7");
END_REGION

REGION Network 2: Acyclic Commands
   RUNG wire#powerrail
      "SLP/SWP331_IOL_Acyclic_Commands_DB"(SystemCommand := "SystemCommand", AcyclicCommandIndex := "AcyclicCommandIndex", AcyclicCommandSubindex := "AcyclicCommandSubindex", AcyclicCommandLength := "AcyclicCommandLength", ParameterValue := "ParameterValue", Send_SystemCmd := "Send_System_Command", Write_AcyclicCommandWithParameter := "Write_CommandWithParameter", Read_AcyclicCommand := "Read_AcyclicCommand", ResetAcyclicBlock := "Reset_Acyclic_Block", SensorStatus =>, ErrorCode =>, Done =>)
   END_RUNG
   // the same network as SCL:
   "SLP/SWP331_IOL_Acyclic_Commands_DB"(SystemCommand := "SystemCommand",   // "SLP/SWP331_IOL_Acyclic_Commands"
                           AcyclicCommandIndex := "AcyclicCommandIndex",
                           AcyclicCommandSubindex := "AcyclicCommandSubindex",
                           AcyclicCommandLength := "AcyclicCommandLength",
                           ParameterValue := "ParameterValue",
                           Send_SystemCmd := "Send_System_Command",
                           Write_AcyclicCommandWithParameter := "Write_CommandWithParameter",
                           Read_AcyclicCommand := "Read_AcyclicCommand",
                           ResetAcyclicBlock := "Reset_Acyclic_Block");
END_REGION
END_FUNCTION

ORGANIZATION_BLOCK "Main"   // OB1, LAD, ProgramCycle
TITLE = "Main Program Sweep (Cycle)"
{ S7_Optimized_Access := 'TRUE' }
VERSION : 0.1
   VAR_INPUT
      Initial_Call : Bool;   // Initial call of this OB
      Remanence : Bool;   // =True, if remanent data are available
   END_VAR
BEGIN

REGION Network 1
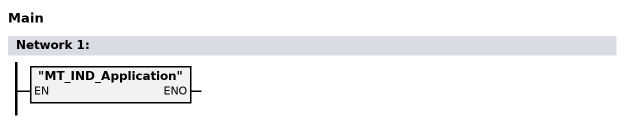
   RUNG wire#powerrail
      "MT_IND_Application"()
   END_RUNG
   // the same network as SCL:
   "MT_IND_Application"();
END_REGION
END_ORGANIZATION_BLOCK

// folder: S7-1200 Basic

FUNCTION_BLOCK "IO_LINK_DEVICE"   // FB50001, SCL
TITLE = IO_LINK_DEVICE
{ S7_Optimized_Access := 'TRUE' }
AUTHOR : SUP_FA
FAMILY : IO-Link
VERSION : 3.0
// Function block to read and write acyclic data on devices with IO-Link used on SIMATIC S7 controllers. (former IO_LINK_CALL)
   VAR_INPUT
      REQ : Bool;   // Request Function / Neuer Auftrag
      ID : Hw_Io;   // Hardwarekennung des IOL-Master Moduls (HW_IO) aus HW-Konfiguration
      CAP : DInt := DINT#0;   // Client Access Point (CAP), bei ET200 immer 227 dez
      RD_WR : Bool;   // Lese und Schreibzugriff auf IO-Link Device 0: Lesen, 1: schreiben
      PORT : Int := INT#0;   // Port/ Kanalnummer an dem das IO-Link Device betrieben wird. (ET200 = 0 .. 4)
      IOL_INDEX : Int := INT#0;   // Adressparameter Index (IO-Link Device) 0..32767 IOL-D, 65535 port functions
      IOL_SUBINDEX : Int := INT#0;   // Adressparameter Subindex (IO-Link Device) 0 ges. Record; 1-255 einz. Parameter
      LEN : Int := INT#0;   // Länge der zu schreibenden Daten (Nettodaten)
   END_VAR
   VAR_OUTPUT
      DONE_VALID : Bool;   // Gültigkeit 0: Daten nicht gültig; 1: Daten gültig
      BUSY : Bool;   // 0: Auftrag abgeschlossen 1: Auftrag in Bearbeitung
      ERROR : Bool;   // Fehler Flag 0: kein Fehler; 1: Abbruch der Funktion mit Fehler
      STATUS : DWord := DWORD#16#0000_0000;   // DP/ PNIO - Fehlerstatus; ERROR Flag = 1 - detaillierter Kommunikationsfehlerstatus
      IOL_STATUS : DWord := DWORD#16#0000_0000;   // IO-Link Fehlerstatus; ERROR Flag = 1 - detaillierte IO-Link Fehlerstatus
      RD_LEN : Int := INT#0;   // Länge des gelesenen Datensatzes (Anzahl Bytes)
   END_VAR
   VAR_IN_OUT
      RECORD_IOL_DATA : Array[0..231] of Byte;   // Datenbereich für LESEN / SCHREIBEN (max. 232 Byte)
   END_VAR
   VAR
      RDREC_Function : RDREC;   // Funktion Datensatz lesen (ehemals SFB52)
      WRREC_Function : WRREC;   // Funktion Datensatz schreiben (ehemals SFB53)
      TP_poll : TP_TIME;   // Pollzeit für "Datensatz lesen"
      TON_monitoring : TON_TIME;   // Überwachungszeit für Aufträge
      rdrec : Struct   // interne Struktur für RDREC
         valid : Bool;   // Function performed
         busy : Bool;   // Function busy
         error : Bool;   // Error flag
         status : DWord;   // Function result/error message
         length : UInt;   // Length of the fetched data record
      END_STRUCT;
      wrrec : Struct   // interne Struktur für WRREC
         length : UInt;   // length of write data record
         done : Bool;   // Function performed
         busy : Bool;   // Function busy
         error : Bool;   // Error flag
         status : DWord;   // Function result/error message
      END_STRUCT;
      read : Struct   // Datenbereich für Lesedaten
         header : Struct
            CALL : Struct   // header for read/write data record
               Extended_Function_Num : Byte := 16#08;   // extended function number (fix coded 08h)
               Port : Byte;   // variable port (user interface) 0...255
               FI_Index : Word := 16#FE4A;   // FI index (fix coded 65098)
            END_STRUCT;
            IOL : Struct   // header for IO-Link
               Control : Byte;   // RD_WR = 0 = read = Control:=0x03 / / RD_WR = 1 = write = Control:=0x02
               Index_HighByte : Byte;   // index of data record 0…32767 (high byte)
               Index_LowByte : Byte;   // index of data record 0…32767 (low byte)
               Subindex : Byte;   // subindex for data record 0...255
            END_STRUCT;
         END_STRUCT;
         data : Array[0..231] of Byte;
      END_STRUCT;
      write : Struct   // Datenbereich für Schreibdaten
         header : Struct
            CALL : Struct   // header for read/write data record
               Extended_Function_Num : Byte := 16#08;   // extended function number (fix coded 08h)
               Port : Byte;   // variable port (user interface) 0...255
               FI_Index : Word := 16#FE4A;   // FI index (fix coded 65098)
            END_STRUCT;
            IOL : Struct   // header for IO-Link
               Control : Byte;   // RD_WR = 0 = read = Control:=0x03 / / RD_WR = 1 = write = Control:=0x02
               Index_HighByte : Byte;   // index of data record 0…32767 (high byte)
               Index_LowByte : Byte;   // index of data record 0…32767 (low byte)
               Subindex : Byte;   // subindex for data record 0...255
            END_STRUCT;
         END_STRUCT;
         data : Array[0..231] of Byte;
      END_STRUCT;
      sequencecontrol : Int := INT#0;   // number of sequence control
      typeofrequest : Int := INT#0;   // type of request (0=Read, 1=Write)
      R_TRIG_REQ : Bool;   // Impuls für neuen Auftrag starten
      R_TRIG_REQ_old : Bool;   // Flankenmerker
      F_TRIG_poll : Bool;   // Impuls für Pollen "Datensatz lesen"
      F_TRIG_poll_old : Bool;   // Flankenmerker
   END_VAR
   VAR_TEMP
      retval : Int;   // Variable für Rückgabewerte von Funktionen
      tmpWORD : Word;   // Datentyp WORD zur temporären Verwendung
      tmpDWORD : DWord;   // Datentyp DWORD zur temporären Verwendung
      tmpINT : Int;   // Datentyp INT zur temporären Verwendung
      i : Int;   // Laufvariable für for-Schleifen
   END_VAR
BEGIN
   (*---------------------------------------------------------------------------------------------------------------------
   SIEMENS AG
   ©Copyright 2017. All Rights Reserved.
   -----------------------------------------------------------------------------------------------------------------------
   Limitation of liability
   This software was developed with largest care. However, the author can not guarantee, that the software runs under
   each version of STEP7 on each PLC flawlessly.
   There is no warranty for the software, to the extent permitted by applicable law. The copyright holder provides the
   software "as is" without warranty of any kind, either expressed or implied, including, but not limited to, the implied
   warranties of merchantability and fitness for a particular purpose. The entire risk as to the quality and performance
   of the software is with you. Should the software prove defective, you assume the cost of all necessary servicing,
   repair or correction. In no event unless required by applicable law will the copyright holder be liable to you for
   damages, including any general, special, incidental or consequential damages arising out of the use or inability to
   use the software (including but not limited to loss of data or data being rendered inaccurate or losses sustained by
   you or third parties or a failure of the software to operate with any other programs), even if such holder or other
   party has been advised of the possibility of such damages.
   Permission to use or copy this software for any purpose is hereby granted without fee, provided the above notices are
   retained on all copies. Permission to modify the code and to distribute modified code is granted, provided the above
   notices are retained, and a notice that the code was modified is included with the above copyright notice.
   -----------------------------------------------------------------------------------------------------------------------
   Functionality provided by this source (short description):
   Function block IO_LINK_DEVICE - used to read and write of acyclic data records on devices with IO-Link.
   Note:
   To read data records, the IO-Link master modules needs to know which data record is required. Therefore it is necessary
   to send at first a request via write data record (only header of 8 byte). As response the IO-Link master module
   will send the required data record.

   Status:     Released (tested)
   File name:  IO_LINK_DEVICE
   System :    SIMATIC S7-1200
   Version :   3.0
   -----------------------------------------------------------------------------------------------------------------------
   Script to be stored on level ... in project (mark appropriate levels with [x] below)
   [ ] External
   [ ] All levels possible
   [x] Project level
   [ ] Controller level
   [ ] Device level
   [ ] Subobject level
   -----------------------------------------------------------------------------------------------------------------------
   Restrictions, known limitations:
   The limitation of 240 byte is based on PROFIBUS DP protocol. With PROFINET IO there wouldn't no limit but because of 
   compatibility reason it wasn't changed.
     - header =   8 byte
     - data   = 232 byte
   -----------------------------------------------------------------------------------------------------------------------
   Requirements, prerequisites, External resources used: nothing
   -----------------------------------------------------------------------------------------------------------------------
   Change log table (latest change is at the bottom OF the list):
   Version Date Changes applied
   V2.0.0 <2013-09-30> First created with TIA Portal V12 SP1
   V2.1.0 <2014-03-14> Upgrade system function 'WRREC' from V1.0 to V1.1 and released for TIA Portal V13
   V3.0.0 <2015-02-28> Upgrade and released for TIA Portal V13 SP1 (without backup/restore master parameter)
   V3.0.2 <2015-07-07> Change of #IOL_INDEX and #Port lower boundry to 0
   V3.0.3 <2017-03-13> Compilation ready for TIA Portal Basic, especially S7-1200 controllers
   ---------------------------------------------------------------------------------------------------------------------*)

   (*---------------------------------------------------------------------------------------------------------------------
   Description of programmed IO-Link error codes
   8000 = time out
   8001 = wrong port
   8002 = wrong index
   8003 = wrong subindex
   8005 = wrong length for write data record
   8006 = wrong length for read data record
   8052 = error during reading data record
   8053 = error during writing data record
   All other codes are coming from a higher level!
   ---------------------------------------------------------------------------------------------------------------------*)

   (*---------------------------------------------------------------------------------------------------------------------
               NEW REQUEST
   ---------------------------------------------------------------------------------------------------------------------*)
   // detection rising edge of "REQ"
   #R_TRIG_REQ := #REQ = TRUE AND #R_TRIG_REQ_old = FALSE;
   #R_TRIG_REQ_old := #REQ = TRUE;

   // start new request if not busy
   IF #R_TRIG_REQ = TRUE AND #sequencecontrol = 0 THEN
       // Freeze record ID and CAP
       #WRREC_Function.ID := #ID;
       #WRREC_Function.INDEX := #CAP;
       #RDREC_Function.ID := #ID;
       #RDREC_Function.INDEX := #CAP;

       // Initialize outputs
       #DONE_VALID := FALSE;
       #BUSY := TRUE;
       #ERROR := FALSE;
       #STATUS := DW#16#00000000;
       #IOL_STATUS := DW#16#00000000;
       #RD_LEN := INT#0;

       // Initialize data area
       #read.header."CALL"."Port" := B#16#0;
       #read.header.IOL.Index_LowByte := B#16#0;
       #read.header.IOL.Index_HighByte := B#16#0;
       #read.header.IOL.Subindex := B#16#0;
       #i := INT#0; // initialize loop counter      
       FOR #i := 0 TO 231 DO
           #write.data[#i] := B#16#0;
           #read.data[#i] := B#16#0;
       END_FOR;

   (*---------------------------------------------------------------------------------------------------------------------
       Setup IO-LINK Call needs a specific header
   ---------------------------------------------------------------------------------------------------------------------*)
   // setup CALL header
   #write.header."CALL".Extended_Function_Num := 16#08;  // extended function number (fix coded 08h)
   #write.header."CALL"."Port" := INT_TO_BYTE(#PORT);  // 1..63 = PORT number, 64..255=reserved
   #write.header."CALL".FI_Index := 65098;  // IOL-Header is following (fix coded 65098)

   // setup IOL header 
   // CONTROL = please see below at BODY
   // INDEX
   #write.header.IOL.Index_LowByte := INT_TO_BYTE(#IOL_INDEX);
   #tmpWORD := INT_TO_WORD(#IOL_INDEX);
   #tmpWORD := SHR(IN := #tmpWORD, N := 8);
   #write.header.IOL.Index_HighByte := WORD_TO_BYTE(#tmpWORD);
   // SUBINDEX
   #write.header.IOL.Subindex := INT_TO_BYTE(#IOL_SUBINDEX);

   // BODY (data max. 232 Byte, Array 0..231 of Byte) 
   IF #RD_WR = TRUE THEN
       // IO-Link write data record requested, copy data from "RECORD_IOL_DATA"
       #write.header.IOL.Control := B#16#02; // CONTROL B#16#02 = write data record
       #wrrec.length := INT_TO_UINT(#LEN) + UINT#8;  // data length header + data = IO-Link write data record
       #typeofrequest := 2; // write data record
       // copy IOL_RECORD_DATA in working area
       #i := INT#0;    // initialize loop counter 
       FOR #i := 0 TO #LEN - 1 DO
           #write.data[#i] := #RECORD_IOL_DATA[#i];
       END_FOR;
   ELSE
       // IO-Link read data record requested
       #write.header.IOL.Control := 16#03;  // CONTROL 16#03 = read data record
       #wrrec.length := UINT#8; // data length only header = IO-Link read data record
       #typeofrequest := 1; // read data record        
   END_IF;
   #sequencecontrol := 1;  // Start sequence
   ELSE
       ;
   END_IF;

   (*---------------------------------------------------------------------------------------------------------------------
               SEQUENCE CONTROL
   ---------------------------------------------------------------------------------------------------------------------*)
   CASE #sequencecontrol OF
       1:  // Check input parameter        
           IF #PORT < INT#0 OR #PORT > INT#63 THEN // PORT (Wrong port address = 0x8001)
               #ERROR := TRUE;
               #IOL_STATUS := DW#16#80010000;
               #sequencecontrol := 99; // aborting function with error
           ELSIF #IOL_INDEX < INT#0 OR #IOL_INDEX > INT#32767 THEN    // INDEX (Wrong index = 0x8002)
               #ERROR := TRUE;
               #IOL_STATUS := DW#16#80020000;
               #sequencecontrol := 99; // aborting function with error
           ELSIF #IOL_SUBINDEX < INT#0 OR #IOL_SUBINDEX > INT#255 THEN    // SUBINDEX (Wrong subindex = 0x8003)
               #ERROR := TRUE;
               #IOL_STATUS := DW#16#80030000;
               #sequencecontrol := 99; // aborting function with error
           ELSIF #typeofrequest = 2 AND (#LEN < 1 OR #LEN > 232) THEN  // LEN (wrong length for write data record = 0x8004)
               #ERROR := TRUE;
               #IOL_STATUS := DW#16#80050000;
               #sequencecontrol := 99; // aborting function with error
           ELSIF #typeofrequest = 1 AND (#LEN < 0 OR #LEN > 232) THEN  // LEN (wrong length for read data record = 0x8005)
               #ERROR := TRUE;
               #IOL_STATUS := DW#16#80060000;
               #sequencecontrol := 99; // aborting function with error
           ELSE    // all input parameter are right
               #sequencecontrol := 2;
           END_IF;

       2:  (*-------------------------------------------------------------------------------------------------------------
           WRREC = Write Data Record
           Note:
           To read data records, the IO-Link master modules needs to know which PORT is required. Therefore it is necessary
           to send at first a request via write data record (header, 8 byte). As response the IO-Link master module will 
           send the required data record.
           -------------------------------------------------------------------------------------------------------------*)
           #WRREC_Function(REQ := TRUE,
                           LEN := #wrrec.length,
                           DONE => #wrrec.done,
                           BUSY => #wrrec.busy,
                           ERROR => #wrrec.error,
                           STATUS => #wrrec.status,
                           RECORD := #write);
           // output status during write data record
           IF #wrrec.busy THEN
               #STATUS := #wrrec.status;
               #IOL_STATUS := DW#16#00020000;  // 0002 = writing in progress 
           ELSIF #wrrec.error THEN
               #tmpDWORD := #wrrec.status AND DW#16#00FFFF00;  // filter status
               IF #tmpDWORD = DW#16#0080C200 THEN    // if resource #BUSY (#STATUS=80C2), then ... 
                   #sequencecontrol := 3;  // ... repeat write data record
               ELSE
                   #ERROR := TRUE;
                   #STATUS := #wrrec.status;   // ... otherwise output error status of "WRREC"
                   #IOL_STATUS := DW#16#80530000;  // ... with note '8053' = error status of "WRREC"
                   #sequencecontrol := 99; // aborting function with error
               END_IF;
           ELSIF #wrrec.done = TRUE THEN   // wait for write data record finish without error
               #TP_poll(IN := TRUE,
                        PT := T#100ms);    // poll for response
               #sequencecontrol := 4;
           ELSE
               ;
           END_IF;

       3:  // repeat write data record because resource was busy
           #WRREC_Function(REQ := FALSE);
           #sequencecontrol := 2;

       4:  // wait and poll for response = Read Data Record (RDREC)
           #WRREC_Function(REQ := FALSE);
           #TP_poll(IN := TRUE,
                    PT := T#100ms);

           // if poll rate executed then start read data record (on falling edge)
           #F_TRIG_poll := #TP_poll.Q = FALSE AND #F_TRIG_poll_old = TRUE;
           #F_TRIG_poll_old := #TP_poll.Q = TRUE;

           // RDREC = Read Data Record
           #RDREC_Function(REQ := #F_TRIG_poll,
                           MLEN := UINT#0, // length = 0 = read all data which are available
                           VALID => #rdrec.valid,
                           BUSY => #rdrec.busy,
                           ERROR => #rdrec.error,
                           STATUS => #rdrec.status,
                           LEN => #rdrec.length,
                           RECORD := #read);
           // output status during read data record
           IF #rdrec.busy THEN
               #STATUS := #rdrec.status;
               #IOL_STATUS := DW#16#00030000; // 16#0003 = reading in progress
           ELSIF #rdrec.error = TRUE THEN
               #tmpDWORD := #rdrec.status AND DW#16#00FFFF00;  // filter status
               IF #tmpDWORD = DW#16#0080C200 THEN  // if resource busy (status=80C2), then ... 
                   #sequencecontrol := 5;  // ... repeat read data record / continue polling
               ELSE
                   #ERROR := TRUE;
                   #STATUS := #rdrec.status;   // ... otherwise output error code of "RDREC"
                   #IOL_STATUS := DW#16#80520000;  // ... with note '8052' = error status of "RDREC"
                   #sequencecontrol := 99; // aborting function with error
               END_IF;
           ELSIF #rdrec.valid THEN
               IF  // check the response wether it matches the request (compare PORT, INDEX and SUBINDEX)
                   (#write.header."CALL"."Port" <> #read.header."CALL"."Port") OR
                   (#write.header.IOL.Index_HighByte <> #read.header.IOL.Index_HighByte) OR
                   (#write.header.IOL.Index_LowByte <> #read.header.IOL.Index_LowByte) OR
                   (#write.header.IOL.Subindex <> #read.header.IOL.Subindex)
               THEN    // read data record don't match the request
                   #ERROR := TRUE;
                   #STATUS := #rdrec.status;
                   #IOL_STATUS := DW#16#70000000;  // output status '7000', no consistent data
                   #sequencecontrol := 99; // aborting function with error
               ELSIF #read.header.IOL.Control = B#16#80 THEN   // check the response for IO-Link errors
                   // State 0x80 = IOL_CALL_RES PDU shows IO-Link error detect
                   #ERROR := TRUE;
                   #STATUS := DW#16#00000000;
                   #IOL_STATUS.%B3 := #read.data[0];   // IO-Link master error code
                   #IOL_STATUS.%B2 := #read.data[1];   // IO-Link master error code
                   #IOL_STATUS.%B1 := #read.data[2];  // IO-Link device error code
                   #IOL_STATUS.%B0 := #read.data[3];  // IO-Link device additional error code

                   #sequencecontrol := 99; // aborting function with error
               ELSE    // read data are valid = output
                   #DONE_VALID := TRUE;
                   #BUSY := FALSE;
                   #ERROR := FALSE;
                   #STATUS := DW#16#00000000;
                   #IOL_STATUS := DW#16#00000000;  // request finished

                   IF #typeofrequest = 1 THEN
                       #RD_LEN := UINT_TO_INT(#rdrec.length - UINT#8);  // device parameter cover header and data,
                       // only data will be output
                       #i := INT#0; // initialize loop counter
                       FOR #i := 0 TO UINT_TO_INT(#rdrec.length - UINT#8 - UINT#1) DO
                           #RECORD_IOL_DATA[#i] := #read.data[#i];
                       END_FOR;
                   ELSE
                       ;
                   END_IF;
                   #sequencecontrol := 98;
               END_IF;
           ELSE
               ;
           END_IF;

       5:  // poll again for response because resource was busy
           #TP_poll(IN := FALSE,
                    PT := T#100ms);
           #RDREC_Function(REQ := FALSE,
                           RECORD := #read);
           #sequencecontrol := 4;  // ... repeat read data record / continue polling   

       98: // request done successfully
           #TP_poll(IN := FALSE,
                    PT := T#100ms);
           #RDREC_Function(REQ := FALSE,
                           RECORD := #read);
           IF #REQ = FALSE THEN
               #DONE_VALID := FALSE;
               #BUSY := FALSE;
               #ERROR := FALSE;
               #RD_LEN := INT#0;
               #STATUS := DW#16#00000000;
               #IOL_STATUS := DW#16#00010000; // ready for new request
               #sequencecontrol := 0;
               #typeofrequest := 0;
           ELSE
               ;
           END_IF;

       99: // Function aborted with error
           #TP_poll(IN := FALSE,
                    PT := T#100ms);
           #WRREC_Function(REQ := FALSE);
           #RDREC_Function(REQ := FALSE,
                           RECORD := #read);
           #DONE_VALID := FALSE;
           #BUSY := FALSE;
           #RD_LEN := INT#0;
           #sequencecontrol := 0;
           #typeofrequest := 0;

       ELSE  // no relevant case, ready for new request
           #WRREC_Function(REQ := FALSE);
           #RDREC_Function(REQ := FALSE,
                           RECORD := #read);
           #TP_poll(IN := FALSE,
                    PT := T#100ms);
           #TON_monitoring(IN := FALSE,
                           PT := T#20s);
           #sequencecontrol := 0;
           #typeofrequest := 0;
   END_CASE;

   (*---------------------------------------------------------------------------------------------------------------------
               MONITORING
   ---------------------------------------------------------------------------------------------------------------------*)
   #TON_monitoring(IN := #sequencecontrol > 0 AND #sequencecontrol < 98,
                   PT := T#20s);
   IF #TON_monitoring.Q THEN
       #ERROR := TRUE;
       #IOL_STATUS := DW#16#80000000; // request time out       
       #sequencecontrol := 99; // aborting function with error
   END_IF;
END_FUNCTION_BLOCK